Fanuc KAREL source: KA00215.KL

PROGRAM KA00215
%NOLOCKGROUP
VAR
  SRC: ARRAY[4] OF XYZWPR
  DST: ARRAY[4] OF XYZWPR
BEGIN
  DST = SRC
END KA00215
